PROGRAM MAIN
VAR
	bCount : BOOL;
	iCounter : INT;
END_VAR

IF bCount THEN
	iCounter := iCounter + 1;
	GVL_SAFETY.bRunStop := TRUE;
END_IF;

END_PROGRAM

(* stored: Version 1.1.0.1, ProductVersion 3.1.4024.12
   POU MAIN: Id {d7652c90-63f4-4e4f-9c9a-cdf0391412f1}, SpecialFunc None *)
